{ attribute 'Name':='TB_Div-Test' }
{ attribute 'Timeout':='t#20s' }
{ attribute 'Owner':='TestOwner' }
{ attribute 'Category':='Math/multiplication and division ' }
FUNCTION_BLOCK FB_TestDiv EXTENDS FB_TestCaseBase
VAR_INPUT
END_VAR
VAR_OUTPUT
END_VAR
VAR
	myFB : SampleLib.FB_Div;    // instance of the function block to be tested
	expectedValue : UINT;       // value to be expected from this test
	result: UINT;				// calculated value, actual result of the function block call
END_VAR

// can of the function block to execute the test: 8 / 2 = 4
myFB(var1:= 8, var2:= 2, result=> result);

// Explicit assignment of the expected value, as the comparison is performed using the “any” data type
expectedValue:=4;

// Check the result against the expected value; if it does not match, the error message passed here is displayed
AssertEqual(anyActual:= result, anyExpected:= expectedValue, sMessage:= 'Division with the FB_Div function block is incorrect!');

// in the event that the result of the comparison matches, confirmation that the test case was successful and that no further tests will be carried out in this function block
Succeed();

//Must be implemented if you want to use fastmode
METHOD CleanUp : BOOL
CleanUp:=true;
END_METHOD

END_FUNCTION_BLOCK

(* stored: Version 1.1.0.1, ProductVersion 3.1.4026.21
   POU FB_TestDiv: Id {b8cf319c-5feb-45d7-908e-09f59f0021f0}, SpecialFunc None
   Method CleanUp: Id {e18a61bd-c4ec-4cd1-b227-251b85e3f0e4} *)
